(* IEC 61131-3 sources: trust-platform/libraries/plant/examples/packaging_machine/src, 3 files *)

(* ---- RejectSequence.st ---- *)
(* Rejects products the inspection marks bad: carries each rejected product to the reject station,
   extends the reject cylinder, and waits for it to retract. A good product passes. *)
USING Plant;

FUNCTION_BLOCK RejectSequence EXTENDS Plant.FB_Sequence
VAR_INPUT
    ProductPresent : BOOL;
    InspectionFailed : BOOL;
    CylinderExtended : BOOL;
    CylinderRetracted : BOOL;
    (* The time a product needs from the sensor to the reject station. *)
    TravelTime : TIME := T#800ms;
END_VAR
VAR_OUTPUT
    RunConveyor : BOOL;
    ExtendCylinder : BOOL;
    Passed : UDINT;
    Rejected : UDINT;
END_VAR
    ExtendCylinder := FALSE;
    IF Execute() THEN
        CASE CurrentStep OF
            0:
                GoTo(Number := 10, Name := 'Wait for a product');
            10:
                Wait(Text := 'Waiting for a product');
                IF ProductPresent THEN
                    IF InspectionFailed THEN
                        GoTo(Number := 20, Name := 'Carry to the reject station');
                    ELSE
                        GoTo(Number := 40, Name := 'Product passes');
                    END_IF;
                END_IF;
            20:
                IF StepTime >= TravelTime THEN
                    GoTo(Number := 30, Name := 'Reject');
                END_IF;
            30:
                ExtendCylinder := TRUE;
                IF CylinderExtended THEN
                    Rejected := Rejected + 1;
                    GoTo(Number := 35, Name := 'Retract');
                ELSE
                    StepTimeout(Limit := T#3s, Text := 'The reject cylinder did not extend');
                END_IF;
            35:
                IF CylinderRetracted THEN
                    GoTo(Number := 10, Name := 'Wait for a product');
                ELSE
                    StepTimeout(Limit := T#3s, Text := 'The reject cylinder did not retract');
                END_IF;
            40:
                IF NOT ProductPresent THEN
                    Passed := Passed + 1;
                    GoTo(Number := 10, Name := 'Wait for a product');
                END_IF;
        END_CASE;
    ELSIF State = E_SequenceState#Stopping THEN
        (* A stop finishes the current product first. *)
        IF CurrentStep = 10 OR CurrentStep = 40 THEN
            StopDone();
        END_IF;
    END_IF;
    RunConveyor := State = E_SequenceState#Running OR State = E_SequenceState#Stopping;
END_FUNCTION_BLOCK

(* ---- Configuration.st ---- *)
CONFIGURATION Packaging
RESOURCE Cpu ON PLC
    TASK Line (INTERVAL := T#10ms, PRIORITY := 1);
    PROGRAM Machine WITH Line : Main;
END_RESOURCE
VAR_CONFIG
    Machine.StartButton AT %IX0.0 : BOOL;
    Machine.StopButton AT %IX0.1 : BOOL;
    Machine.ProductSensor AT %IX0.2 : BOOL;
    Machine.InspectionFailed AT %IX0.3 : BOOL;
    Machine.ConveyorRunning AT %IX0.4 : BOOL;
    Machine.ConveyorTrip AT %IX0.5 : BOOL;
    Machine.CylinderExtendedSensor AT %IX0.6 : BOOL;
    Machine.CylinderRetractedSensor AT %IX0.7 : BOOL;
    Machine.ConveyorRun AT %QX0.0 : BOOL;
    Machine.RejectValve AT %QX0.1 : BOOL;
END_VAR
END_CONFIGURATION

(* ---- Main.st ---- *)
(* Packaging line: an infeed conveyor carries products past a product sensor and the inspection
   result; RejectSequence pushes bad products off with a single-acting reject cylinder. *)
USING Plant;

PROGRAM Main
VAR
    (* Hardware signals, mapped to I/O in Configuration.st. *)
    StartButton : BOOL;
    StopButton : BOOL;
    ProductSensor : BOOL;
    InspectionFailed : BOOL;
    ConveyorRunning : BOOL;
    ConveyorTrip : BOOL;
    CylinderExtendedSensor : BOOL;
    CylinderRetractedSensor : BOOL;
    ConveyorRun : BOOL;
    RejectValve : BOOL;

    Product : Plant.FB_DigitalInput := (Debounce := T#20ms);
    Conveyor : Plant.FB_Conveyor;
    Reject : Plant.FB_Cylinder := (ExtendTimeout := T#1s, RetractTimeout := T#1s);
    Line : RejectSequence;
    StartEdge : R_TRIG;
    StopEdge : R_TRIG;
END_VAR
    Product(Input := ProductSensor);
    StartEdge(CLK := StartButton);
    StopEdge(CLK := StopButton);
    IF StartEdge.Q THEN
        Line.Start();
    END_IF;
    IF StopEdge.Q THEN
        Line.Stop();
    END_IF;
    Line(ProductPresent := Product.Value, InspectionFailed := InspectionFailed,
        CylinderExtended := Reject.Extended, CylinderRetracted := Reject.Retracted);
    Conveyor(AutoRun := Line.RunConveyor, RunningFeedback := ConveyorRunning, Trip := ConveyorTrip);
    Reject(AutoExtend := Line.ExtendCylinder, ExtendedSensor := CylinderExtendedSensor,
        RetractedSensor := CylinderRetractedSensor);
    ConveyorRun := Conveyor.RunCommand;
    RejectValve := Reject.ExtendCommand;
END_PROGRAM
